// TIA Portal V20 export
FUNCTION "Block_2" : Void   // FC1, LAD
{ S7_Optimized_Access := 'TRUE' }
// stored: SetENOAutomatically false
BEGIN

REGION Network 1
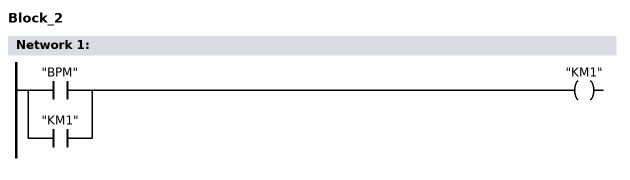
   RUNG wire#powerrail
      Contact( "BPM" )
      wire#w1
      Coil( "KM1" )
   END_RUNG
   RUNG wire#powerrail
      Contact( "KM1" )
   END_RUNG wire#w1
   // the same network as SCL:
   "KM1" := "BPM" OR "KM1";
END_REGION
END_FUNCTION
